// TIA Portal V21 export
// export: Created 2026-11-18T04:37:20.4003739Z, ExportSetting WithDefaults, DisplayName Totally Integrated Automation Portal, DisplayVersion V21, DisplayName STEP 7 Professional, DisplayVersion V21, DisplayName STEP 7 Safety, DisplayVersion V21, DisplayName Tech WebApplication, DisplayVersion V21, DisplayName WinCC Basic/Comfort/Advanced, DisplayVersion V21
TagTable "Default tag table"
  Tag_ScreenNumber : UInt  (1 s)
